// Réponse de I_Object.Start (docs/04 § 5)
{attribute 'qualified_only'}
{attribute 'strict'}
TYPE E_StartResult :
(
    Accepted := 0,
    Busy := 1,
    NotReady := 2,
    UnknownAction := 3,
    BadParam := 4,
    Interlocked := 5,
    Disabled := 6,
    ManualOnly := 7,
    NotConfigured := 8
) USINT;
END_TYPE

(* stored: Version 1.1.0.1, ProductVersion 3.1.4024.12
   DUT E_StartResult: Id {771fb800-cabc-569a-9b9b-c19fa2033346} *)
